Omron CX-Programmer project  (CX-Programmer ?)

# PLC :  

## Global symbols (name address type ; comment)
W4.01 BOOL  ; Лифт №1 РЕЛЕ ВКЛ питание
W5.01 BOOL  ; Лифт №1 Реле выкл Питание
BLINK_L1 BLINK
DOWN W1.03 BOOL
DOWN_stop W0.03 BOOL
HOME_L1 W0.08 BOOL  ; Лифт откальброван
L1_DOWN W0.00 BOOL
L1_UP W0.01 BOOL
L2_DOWN W0.04 BOOL
L2_DOWN_stop W0.07 BOOL
L2_UP W0.05 BOOL
L2_UP_stop W0.06 BOOL
ON W1.00 BOOL
UP W1.02 BOOL
UP_stop W0.02 BOOL

## Program Probe (cyclic task 0)
Local symbols
BLINK_1_OUT W1.01 BOOL
L1_Key_start 0.08 BOOL  ; $?St$Bk?_#[314] / Лифт №1 Кнопка "Старт"$?St$Bk?_#[314]
L1_Key_stop 0.09 BOOL  ; $?St$Bk?_#[315] / Лифт №1 Кнопка "Стоп"$?St$Bk?_#[315]
L1_Lamp_start 3.06 BOOL  ; Лифт №1 Лампа Старт
L1_in_N_limit 1.06 BOOL  ; Лифт №1 Нижний аварийный концевик
L1_in_P_limit 1.07 BOOL  ; Лифт №1 Верхний аварийный концевик
L1_out_Down 4.08 BOOL  ; Лифт №1 Реле ВКЛ движение вниз
L1_out_Drag 4.12 BOOL  ; Лифт №1 Реле отключение тормоза
L1_out_Up 4.10 BOOL  ; Лифт №1 Реле ВКЛ движение вверх
L1_out_powerON 4.14 BOOL  ; Лифт №1 Реле ВКЛ питание

### Section Main

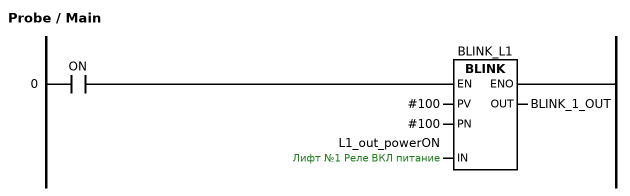
; rung 0
LD ON
CALL BLINK_L1 : BLINK (PV := #100, PN := #100, IN := L1_out_powerON, OUT => BLINK_1_OUT)  ; Лифт №1 Реле ВКЛ питание
; rung 1
END

## Function block BLINK
VAR_INPUT
  PV : INT;
  PN : INT;
  IN : BOOL;
END_VAR
VAR_OUTPUT
  OUT : BOOL;
END_VAR
VAR
  TIMER_1 : TIMER;
  TIMER_2 : TIMER;
  ON : BOOL;
END_VAR

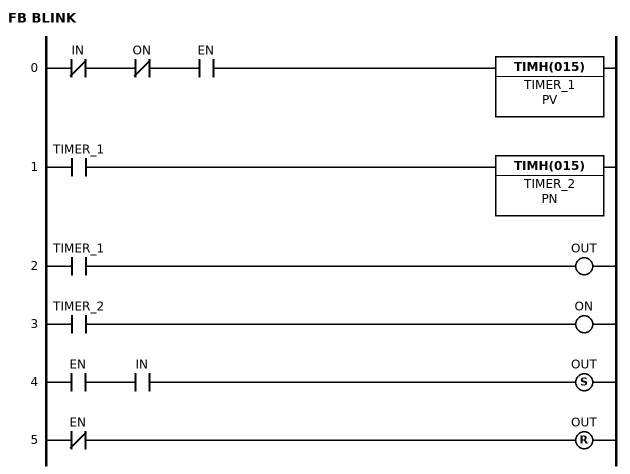
; rung 0
LDNOT IN
ANDNOT ON
AND EN
TIMH(015) TIMER_1 PV
; rung 1
LD TIMER_1
TIMH(015) TIMER_2 PN
; rung 2
LD TIMER_1
OUT OUT
; rung 3
LD TIMER_2
OUT ON
; rung 4
LD EN
AND IN
SET OUT
; rung 5
LDNOT EN
RSET OUT